(*
SPDX-License-Identifier: MIT
License: https://opensource.org/license/mit
*)

(*!
<summary>Owns one single-cycle regression test.</summary>
<description>
Owns persistent child storage and fixed parent associations. Use in one task without reentry.
Children is borrowed and must not be modified by application code. Constructor callbacks are not used.
</description>
*)

{attribute 'no_assign'}
{attribute 'no_explicit_call' := 'do not call this function block directly'}
FUNCTION_BLOCK SingleChildTestGroup EXTENDS TOF_Testing.TestGroup<1>
VAR_STAT
	//! <summary>Class name shared by all instances of this function block.</summary>
	{attribute 'hide'}
	_ClassName : STRING := __POUNAME();
END_VAR
VAR
	{attribute 'hide'}
	{attribute 'init_namespace'}
	_NamespaceName : STRING;
END_VAR
VAR_OUTPUT
	//! <summary>Owned leaf exposed for regression observations and scenario selection.</summary>
	Child : TestingProbe(name := "Owned leaf", parent := THIS^);
END_VAR
VAR
	_Children : ARRAY [0.._ChildCount - 1] OF TOF_Testing.ITestElement :=
	[
		Child
	];
END_VAR

//! <summary>Borrows the concrete class name for the lifetime of this instance; callers must not modify it.</summary>
{attribute 'monitoring' := 'call'}
PROPERTY ClassName : REFERENCE TO STRING
GET
ClassName REF= _ClassName;
END_GET
END_PROPERTY

//! <summary>Borrows the compiler-initialized namespace; callers must not modify the returned reference.</summary>
{attribute 'monitoring' := 'call'}
PROPERTY NamespaceName : REFERENCE TO STRING
GET
NamespaceName REF= _NamespaceName;
END_GET
END_PROPERTY

//! <summary>Reports the complete concrete instance size, excluding separately allocated storage.</summary>
{attribute 'monitoring' := 'call'}
PROPERTY SelfSize : ULINT
GET
SelfSize := XSIZEOF(THIS^);
END_GET
END_PROPERTY

//! <summary>Borrows the fixed array of this concrete group; do not modify it.</summary>
{attribute 'monitoring' := 'call'}
PROPERTY Children : REFERENCE TO ARRAY [0.._ChildCount - 1] OF TOF_Testing.ITestElement
GET
Children REF= _Children;
END_GET
END_PROPERTY

END_FUNCTION_BLOCK

(* stored: Version 1.1.0.1
   POU SingleChildTestGroup: Id {08bf5c2e-1597-4e8a-a0fa-72b8815c4d37}, SpecialFunc None
   Property ClassName: Id {ecb4d9f9-dc49-4312-85f4-41522a872232}
   Get Get: Id {60cdf768-79d5-46e6-84b8-0443346de98d}
   Property NamespaceName: Id {9317d75c-8ab9-4f43-8f5c-5e8fd57d7d67}
   Get Get: Id {7333a108-7a42-4245-9054-eb08efd1f200}
   Property SelfSize: Id {786a3593-d457-49e1-8cb5-cb957090e0ed}
   Get Get: Id {bc944358-bae1-4276-a49c-d651ae4c8569}
   Property Children: Id {2dcc93e6-a44b-4d17-8ecb-e3286b223353}
   Get Get: Id {d096cd8e-b9fa-4f0e-b845-538a1081d88c} *)
